Staubli VAL3: paraStart.pgx

program paraStart(num x_nPoint)
begin

  //  call trajectory:getPointPara(sTrajItem,x_nPoint,nMoveType,nParaSpeed,nParaAccel,nParaBlend,nParaPercent,sComment,bSafePoint,sBlendType,nTRSF,sTRSF)
  //  switch nMoveType
  //    case 0
  //      sParaType="POINT"
  //    break
  //    case 1
  //      sParaType="JOINT"
  //    break
  //  endSwitch

  call trajectory:getPointPara(sTrajItem,x_nPoint,nMoveType,nParaSpeed,nParaAccel,nParaBlend,nParaPercent,sComment,bSafePoint,sBlendType,nTRSF,sTRSF)
  switch nMoveType
    case 1
      bShow2Point=false
      resize(sParaPointType,1,2)
      sParaPointType[0]="POINT"
      sParaPointType[1]="JOINT"
      sParaType="POINT"
    break
    case 0
      bShow2Point=false
      resize(sParaPointType,1,2)
      sParaPointType[0]="POINT"
      sParaPointType[1]="JOINT"
      sParaType="JOINT"
    break
    case 2
      bShow2Point=true
      resize(sParaPointType,1,1)
      sParaPointType[0]="CIRCLE"
      sParaType="CIRCLE"
    break
  endSwitch
end
